Fanuc KAREL source: ko00065.KL

-- PROVISIONAL review KL for V770-1; original PC SHA256 4cd6650e851d74e55e20e12debaef8217dd110a927eb5518279739e73bb1a1b0
-- Incomplete behavior may be omitted. Consult companion uncertainty JSON. Do not deploy.
PROGRAM KO00065
%NOLOCKGROUP
BEGIN
  -- UNRESOLVED_PC offsets 5-12; opcodes 9D,23
  -- UNRESOLVED_PC offsets 17-63; opcodes 27,22,1C,22,1C,22,31,7E,4A
  -- UNRESOLVED_PC offsets 68-72; opcodes 7F
END KO00065
